(* IEC 61131-3 sources: IRIS-Project/LASAL CONTROL SOFTWARE/LasalProject_2025_09_12/Runtime/%LASALAPPDATA%/Runtime/Library/Loader/Source/code (part 4) *)

Find_sRam_I_END

END_FUNCTION // Find_sRam_I
#endif

FUNCTION GLOBAL Find_sRamEx
VAR_INPUT
	CRC32		: UDINT;
  bDontAdd : BOOL;
END_VAR
VAR_OUTPUT
	pRamAdr			: ^XramCell;
END_VAR
VAR
	pRamAdr_Kopie	: ^XramCell;
	udAllocated : UDINT;
	udLength : UDINT;
	RelAdress		: UDINT;
	pData : ^USINT;
	pData_Kopie : ^USINT;
	errCode : DINT;
	rc : DINT;
END_VAR

	IF fReorgSram THEN
		rc := LoadSramKopie(#errCode, 0, 0);
		IF rc <> 0 THEN
			// das Laden de SRAM Kopie hat nicht funktioniert
			fReorgSram := 0;
			DEBUGLOG2("%010d LoadSramKopie failed, rc=%d, errCode = 0x%X" , rc$UDINT, errCode$UDINT);
		END_IF;
	END_IF;

	IF fReorgSram THEN
		// in der Kopie suchen
		pRamAdr := Find_sRam_I(_S_RAM_Hptr_Kopie, CRC32);
	ELSE
		// im SRAM suchen
		pRamAdr := Find_sRam_I(_S_RAM_Hptr, CRC32);
	END_IF;

	IF pRamAdr = NIL THEN
		// nicht gefunden (weder im SRAM noch in der Kopie), neue Zelle anlegen
    if(bDontAdd = FALSE) then
  		nbrOfCells_notFound += 1;
  		pRamAdr := Add_sRam_I(CRC32);
    end_if;

	ELSIF fReorgSram THEN
		// in der Kopie gefunden, Zelle aus der Kopie ins SRAM kopieren
		nbrOfCells_foundInCopy += 1;

		pRamAdr_Kopie := pRamAdr;
		pRamAdr := Add_sRam_I(CRC32);
		IF pRamAdr THEN
			IF (pRamAdr_Kopie^.udType AND 16#3C000000) = IsXram THEN
				// RAMEX Zelle
 		     	udLength := pRamAdr_Kopie^.udData shr 16;
				// wenn die Länge der Daten > 0 ist, dann muss das RAMEX Objekt mit
				// den Daten aus der Kopie vorgeladen und für gültig erklärt werden
				IF udLength > 0 THEN
				 	RelAdress$UDINT:= (SRAM_GetMemory(udLength))$UDINT;
				 	// --- Speicher ist zugewiesen worden --
				 	If RelAdress <> 0 THEN
				   		GET_USED_S_RAM();
				   		udAllocated		      := SRAM_GET_ALLOCATED(udLength);
			  	   		pRAMadr^.udData$UDINT := (udLength shl 16) or (udAllocated and 16#ffff);
				   		pRAMadr^.udType 	  := RelAdress;
				   		pData				  := _S_RAM_Hptr^.DataStart+RelAdress;
				   		pData_Kopie			  := _S_RAM_Hptr_Kopie^.DataStart+(pRamAdr_Kopie^.udType and 16#00FF_ffff);
				   		_memcpy(pData, pData_Kopie, udLength);   // Speicher aus dem Inhalt aus der Kopie vorladen
		           		MakeRamExChk(pRAMadr);

				 	// -- Kein speicher verfügbar !!
				 	ELSE

						pRAMadr := NIL;

				 	END_IF;
				ELSE
	           		MakeRamExChk(pRAMadr);
				END_IF;
			ELSE
				// RAM Zelle
				pRamAdr^.udData := pRamAdr_Kopie^.udData;
				pRamAdr^.udChk := pRamAdr^.udData + CRC32;
				pRamAdr^.udType := 16#C0000000;    // ganz am ende machen wir uns gültig !
			END_IF;
		END_IF;
	ELSE
		nbrOfCells_foundInSram += 1;
	END_IF;

END_FUNCTION

FUNCTION GLOBAL Find_sRam
VAR_INPUT
	CRC32		: UDINT;
END_VAR
VAR_OUTPUT
	pRamAdr			: ^XramCell;
END_VAR

  pRamAdr := Find_sRamEx(CRC32, FALSE);

END_FUNCTION

////////////////////////////////////////////////////////////////////
//
//  Die IDEE:
//
//  LDRMEM => STRUCT
//
//  +----+-------------------------------+------------------------
//  |INFO| Allocation Table:             |
//  |MAT |   einzele Bits geben benutze  |   DATEN in 16-Byte Blöcken
//  |    |   Blöcke an                   |
//  +----+-------------------------------+------------------------
//
//  Allocation Table:
//  - jedes Bit kennzeichnet einen Block in den Daten
//  - ein 1er im Bit sagt aus, daß der entsprechende Block in den Daten frei ist
//  - das MSB zeigt auf den Block mit der höheren Adresse
//
//
////////////////////////////////////////////////////////////////////

FUNCTION SRAM_GetMemoryEx
VAR_INPUT
   length0  : UDINT;
   pGotMemory : ^BOOL;  // Da beim Returnwert 0 nicht unterschieden werden kann, ob
                        // der Offset 0 gemeint ist oder Out-Of-Memory, wird mit diesem
                        // Flag angezeigt, ob Speicher allokiert werden konnte.
END_VAR
VAR_OUTPUT
   ret0 : ^USINT;
END_VAR
VAR
   allocblocknum : UDINT;
   allocblocknumorg : UDINT;
   matsize  : UDINT;
   actblockcount : UDINT;
   actblocknum : UDINT;
   fbptr:^usint;
   startptr:^usint;
   fb, xfb : usint;
   bitcounter:usint;
   start:usint;
   startbit:usint;
   bytecounter:udint;
END_VAR

  pGotMemory^ := FALSE;
  ret0 := NIL; 	//#FA16122003
  if length0 = 0 then
    ret0 := NIL;
    return;
  end_if;

  allocblocknum := ((length0-1) / pLdrmem^.blocksize)+1; // Anzahl der erforderlichen Blöcke
  allocblocknumorg := allocblocknum;
  matsize := pLdrmem^.matsize; // Größe der MAT in Bytes
  actblockcount := 0;
  fbptr := #pLdrmem^.mat[0];
  fb := fbptr^;
  start := 1; // 1=suche ersten freien Block, 0=freier wurde Block gefunden
  bytecounter := 0;

  // Schleife, in der die MAT nach einem zusammengehörenden Bereich mit freien
  // Blöcken (=gesetzten Bits) durchsucht wird.
  while matsize do
    fb := fbptr^;
    if fb then
      // das aktuelle Byte in der MAT ist <>0, d.h. manche Blöcke sind frei
      if start = 0 then
        bytecounter += 1;
      end_if;

      // alle Bits des Bytes fb durchgehen
      bitcounter := 0;
      while bitcounter < 8 do
        xfb := fb and 1;
        fb  := fb shr 1;
        if xfb then
          // wir sind innerhalb des Bytes auf einen freien Block gestoßen
          if start then
            // es handelt sich um den ersten freien Block
            start := 0;
            startptr := fbptr;
            startbit := bitcounter;
            allocblocknum := allocblocknumorg;
            actblocknum := actblockcount;
            bytecounter := 0;
          end_if;
          allocblocknum -= 1;
          if allocblocknum = 0 then
            // es wurde ein zusammenhängender Bereich freier Blöcke gefunden
            ret0 := NIL + ((actblocknum * 8) + startbit) * pLdrmem^.blocksize;
            pGotMemory^ := TRUE;

            // es müssen jetzt noch die Bits in der MAT auf den Wert 'belegt'(=0) geändert werden
            if bytecounter = 0 then   // startbit and endbit same byte
              // auf fb wird jetzt eine Maske geschrieben, mit der dann die Bits auf 0 ausmaskiert werden können
              if startbit = bitcounter then   // only a block of 16 byte
                fb := not (1 shl bitcounter);
              else
                bitcounter := 7 - bitcounter;
                fb := ((16#FF shr startbit) and 16#FF) shl startbit; // Bits rechts von startbit werden auf 0 gesetzt
                fb := ((fb shl bitcounter) and 16#FF) shr bitcounter; // Bits links von bitcounter werden auf 0 gesetzt
                fb := not fb; // Wert invertieren, damit er als UND-Maske verwendet werden kann
              end_if;
              startptr^ := startptr^ and fb; // Bits mit der Maske auf 0 ausmaskieren
            else // 1 byte between start and end
              fb := ((16#FF shr startbit) and 16#FF) shl startbit; // Bits rechts von startbit werden auf 0 gesetzt
              fb := not fb; // Wert invertieren, damit er als UND-Maske verwendet werden kann
              startptr^ := startptr^ and fb; // Bits mit der Maske auf 0 ausmaskieren
              startptr += 1;
              if bytecounter then
                bytecounter -= 1;
                // die Bytes zwischen dem ersten und letzten werden zur Gänze auf 0 gesetzt
                while bytecounter do
                  startptr^ := 0;
                  startptr += 1;
                  bytecounter -= 1;
                end_while;
              end_if;
              bitcounter := 7 - bitcounter;
              fb := ((16#FF shl bitcounter) and 16#FF) shr bitcounter;// Bits links von bitcounter werden auf 0 gesetzt
              fb := not fb; // Wert invertieren, damit er als UND-Maske verwendet werden kann
              startptr^ := startptr^ and fb; // Bits mit der Maske auf 0 ausmaskieren
            end_if;

            // Fertig !
            return;

          end_if;
        else
          // wir sind innerhalb des Bytes auf einen belegten Block gestoßen
          start := 1;
        end_if;
        bitcounter += 1;
      end_while;
    else // if fb
      // das aktuelle Byte in der MAT ist 0, d.h. alle Blöcke sind belegt
      start := 1;
    end_if;
    actblockcount += 1;
    fbptr += 1;
    matsize -= 1;
  end_while;

END_FUNCTION

FUNCTION GLOBAL SRAM_GetMemory
VAR_INPUT
   length0  : UDINT;
END_VAR
VAR_OUTPUT
   ret0 : ^USINT;
END_VAR
VAR
	gotMemory : BOOL;
END_VAR

  ret0 := SRAM_GetMemoryEx(length0, #gotMemory);

END_FUNCTION

//---------------------------------------------
// Speicher Belegen
//---------------------------------------------
// es werden immer ganze blöcke vergeben
// -> Raladdr0 = Startadresse im s-Ram
// ->  length0 = Speicherlänge
//     #FA vorsicht die length hat 2 teile byte0/1 ist die allocated length
//                                         byte2/3 ist die used length
//										   also ein mask ist wichtig

// Wenn in length0 das oberste Bit gesetzt ist, dann wird vor dem Belegen geprüft,
// ob der gesamte Bereich frei ist. Wenn er nicht frei ist, dann wird auch nichts
// belegt.

//<-- 0 wenn ok

// diese Funktion wird nur beim Start verwendet um die bereits belegten RAMZellen zu markieren
// in Version alt 1 Bit sind 16 Byte
// in Version neu 1 Bit sind  4 Byte (der Rest der INFO steht im File beim C-IPC)
// abfrage über version die in den oberen 16 Bit von DataValid steht

FUNCTION SRAM_MarkMemory2
VAR_INPUT
   reladdr0 :^usint;
   length0  : UDINT;
END_VAR
VAR_OUTPUT
   ret0 : DINT;
END_VAR

    IF length0 AND 16#80000000 THEN
        // prüfen, ob der gesamte Bereich belegt ist
        length0 -= 16#80000000;
        ret0 := SRAM_FreeMarkMemory(reladdr0$UDINT, length0, 0, TRUE);
        IF ret0 <> 0 THEN
            RETURN;
        END_IF;
    END_IF;

    ret0 := SRAM_FreeMarkMemory(reladdr0$UDINT, length0, 1(*mark*), FALSE);

END_FUNCTION

#ifdef _LSL_TARGETARCH_ARM
FUNCTION GLOBAL SRAM_MarkMemory
VAR_INPUT
   reladdr0 :^usint;
   length0  : UDINT;
END_VAR
VAR_OUTPUT
   ret0 : DINT;
END_VAR

  ret0 := SRAM_MarkMemory2(reladdr0, length0);

END_FUNCTION
#else
FUNCTION AWL GLOBAL SRAM_MarkMemory
VAR_INPUT
   reladdr0 :^usint;
   length0  : UDINT;
END_VAR
VAR_OUTPUT
   ret0 : DINT;
END_VAR
    PUSHAD

    push      eax         //Result
    push.d    length0
    push.d    reladdr0

    call      SRAM_MarkMemory2

    add.esp   8
    pop.d     ret0        //Result

	POPAD

END_FUNCTION
#endif

#ifdef _LSL_TARGETARCH_ARM
FUNCTION GLOBAL SRAM_UnmarkMemory
VAR_INPUT
   reladdr0 :^usint;
   length0  : UDINT;
END_VAR
VAR_OUTPUT
   ret0 : DINT;
END_VAR

  ret0 := SRAM_FreeMarkMemory(reladdr0$UDINT, length0, 0(*0=Free Memory*), 0(*FALSE:ändern*));

END_FUNCTION
#else
FUNCTION AWL GLOBAL SRAM_UnmarkMemory
VAR_INPUT
   reladdr0 :^usint;
   length0  : UDINT;
END_VAR
VAR_OUTPUT
   ret0 : DINT;
END_VAR
    PUSHAD

    //#SR 16.12.2005
    push      eax         //Result
    push.d    0           //check
    push.d    0           //for unmark memory
    push.d    length0
    push.d    reladdr0

    call      SRAM_FreeMarkMemory

    add.esp   16
    pop.d     ret0        //Result

	POPAD

END_FUNCTION
#endif

//-------------------------------------------
//--- S-Ram Speicherverwaltung Initialisieren
//-------------------------------------------

// Hat a.m geprüft

FUNCTION GLOBAL SRAM_Startup
VAR_INPUT
   length0  : UDINT;
   clear0   : UDINT;
END_VAR
VAR_OUTPUT
   ret0 : DINT;
END_VAR
VAR
   matsize  : UDINT;
   memlength  : UDINT;
END_VAR

   ret0 := -1; // desciptior fehlerhaft, nichts gibts für die ramexerei

   // Größe der MAT ermitteln
   if !!isRamfileDatUsed | ((_S_RAM_Hptr^.DataValid SHR 16) < 2)  then
    matsize   := length0 / (CST_SRAM_BLOCKSIZE * 8); // anzahl der BitMarker
    memlength := matsize * (CST_SRAM_BLOCKSIZE * 8);
   else
    matsize   := 4 * length0 / (CST_SRAM_BLOCKSIZE * 8); // anzahl der BitMarker
    memlength := matsize * (CST_SRAM_BLOCKSIZE * 8) / 4;
   end_if;

   IF pLdrmem = NIL THEN
    // MAT neu allokieren
	// pr:
	//	In der Funktion SRAM_ClearMAT wird um ein DWORD mehr als matsize initialisiert,
	//  daher müssen 4 Bytes zusätlich allokiert werden. Den Grund für die zusätzlichen
	//	4 Bytes kenne ich nicht.
   	pLdrmem := _alloc_resize_LDR(MAT_INFO_TYPE.mat + matsize + 4)$^MAT_INFO_TYPE;
   ELSIF pLdrmem^.matsize <> matsize THEN
    // Größe der MAT ändern
   	pLdrmem := _realloc_LDR(pLdrmem, MAT_INFO_TYPE.mat + matsize + 4)$^MAT_INFO_TYPE;
   END_IF;

   IF pLdrmem = NIL THEN
    ret0 := -1;
    RETURN;
   END_IF;

   pLdrmem^.memlength := memlength;
   pLdrmem^.matsize   := matsize;
   if !!isRamfileDatUsed | ((_S_RAM_Hptr^.DataValid SHR 16) < 2)  then
	pLdrmem^.blocksize := CST_SRAM_BLOCKSIZE;
   else
	pLdrmem^.blocksize := CST_SRAM_BLOCKSIZE_NEW;
   end_if;

   if clear0 then
    SRAM_ClearMAT();
   end_if;

   ret0 := 0; // alles ist gut, daher probieren mal eine kleine ramexerei
END_FUNCTION

//---------------------------------------------
// -- ALLE Blockmarker mit 1 auf "leer" setzen
//---------------------------------------------
#ifdef _LSL_TARGETARCH_ARM
FUNCTION GLOBAL SRAM_ClearMAT

  _memset(#pLdrmem^.mat[0], 16#ff, pLdrmem^.matsize);

END_FUNCTION
#else
FUNCTION AWL GLOBAL SRAM_ClearMAT

		l.ecx		pLdrmem
   		l.ecx		(ecx + MAT_INFO_TYPE.matsize)
		shr.ecx		2				// /4
		jecxz		SRAM_ClearMATRet

		// pr: wozu das ???
		// ** Fehler IPC 300 **     // es wird mehr eigetragen wie vorhandener speicher
		inc			ecx				// wegen IPC 300 sonst werden die Daten nicht gespeichert

		l.edi		pLdrmem
		add.edi		MAT_INFO_TYPE.mat
		l.eax		16#ffffffff
		rep
		stosd
SRAM_ClearMATRet
END_FUNCTION
#endif

//-----------------------------------
// Liefert Die Belegte Speichergrösse (bezogen auf speicherstart)
//-----------------------------------
FUNCTION GLOBAL SRAM_GetLastAddr
VAR_OUTPUT
   ret0 : UDINT;
END_VAR
VAR
   Lng: UDINT;
   size:udint;
   Muster : BSINT;
   fbptr : ^bsint;
END_VAR
   fbptr := #pLdrmem^.mat[pLdrmem^.matsize-1];  // in letzet eintrag im array

   Lng    := pLdrmem^.memlength;				// beginn bei voller belegung
   size   := pLdrmem^.matsize;

   while size do
      if fbptr^ <> 16#FF then     			// erster freier platz wenn nicht auf FF
		 Muster:=fbptr^ $bsint;
		 While Muster do
           Lng-=pLdrmem^.blocksize;
		   muster := muster SHL 1;
		 end_while;
		 Goto  LastAdrEnde;

      end_if;
      fbptr -= 1;
	  size -= 1;
	  Lng-= pLdrmem^.blocksize*8;
   end_while;

LastAdrEnde:
   ret0 := Lng;
END_FUNCTION

(*
    Markiert im Sram in der MAT einen Bereich als frei oder belegt oder
    prüft ob der Bereich vollständig frei oder vollständig belegt ist.
*)
FUNCTION SRAM_FreeMarkMemory
VAR_INPUT
    reladdr0 : UDINT;
    length0  : UDINT;
    mode0    : UDINT;        //0=Free Memory, 1=Mark Memory
    check0   : BOOL;         //FALSE:ändern, TRUE:nur prüfen
END_VAR
VAR_OUTPUT
    ret0 : DINT;
END_VAR
VAR
    startBit : UDINT;
    endBit : UDINT;
    curBit : UDINT;
    ofs : UDINT;
    pMat : ^USINT;
    matVal : USINT;
END_VAR

    ret0 := 0;

    IF ((reladdr0 + length0) > pLdrmem^.memlength) | (length0 = 0) THEN
        // Der angegebene Bereich liegt ausserhalb der Grenzen oder die Länge ist 0 -> Fehler zurückgeben
        ret0 := -1;
        RETURN;
    END_IF;

    startBit := reladdr0 / pLdrmem^.blocksize;
    endBit := (reladdr0 + length0 - 1) / pLdrmem^.blocksize;
    IF mode0 = 0 THEN
        matVal := 0xFF;
    ELSE
        matVal := 0x00;
    END_IF;

    curBit := startBit;
    pMat := #pLdrmem^.mat[curBit / 8];
    WHILE curBit <= endBit DO
        ofs := curBit MOD 8;
        IF (ofs = 0) & ((endBit - curBit) >= 8) THEN
            // Wir befinden uns auf einer Byte-Grenze daher können alle 8 Bits
            // des MAT-Bytes auf einmal behandelt werden.
            IF check0 THEN
                // nur prüfen
                IF pMat^ <> matVal THEN
                    ret0 := -1;
                    RETURN;
                END_IF;
            ELSE
                // ändern
                pMat^ := matVal;
            END_IF;

            curBit += 8;
            pMat += 1;
        ELSE
            // Wir befinden uns mitten im Byte. Die Bits müssen einzeln behandelt werden.
            IF check0 THEN
                // nur prüfen
                IF mode0 = 0 THEN
                    IF (pMat^ AND (1 SHL ofs)$USINT) = 0 THEN
                        ret0 := -1;
                        RETURN;
                    END_IF;
                ELSE
                    IF (pMat^ AND (1 SHL ofs)$USINT) <> 0 THEN
                        ret0 := -1;
                        RETURN;
                    END_IF;
                END_IF;
            ELSE
                // ändern
                IF mode0 = 0 THEN
                    pMat^ := pMat^ OR (1 SHL ofs)$USINT;
                ELSE
                    pMat^ := pMat^ AND NOT (1 SHL ofs)$USINT;
                END_IF;
            END_IF;

            curBit += 1;
            IF (curBit MOD 8) = 0 THEN
                pMat += 1;
            END_IF;
        END_IF;
    END_WHILE;

END_FUNCTION

#ifdef LDR_RETSVR
FUNCTION GLOBAL GetNbrNotFound
VAR_OUTPUT
  ret0 : udint;
END_VAR

  ret0 := nbrOfCells_notFound;

END_FUNCTION

// ein neues File muss erstellt werden
FUNCTION NewRetainSvrFile
	VAR_INPUT
		usProbe 	: usint;
	END_VAR
  VAR_OUTPUT
    ok : dint;
  END_VAR
  var
    pRead : ^MRAM_DESCR;
    pData : ^MRAM_DESCR;
  end_var

  // Schreib-/Lesebuffer
  pData := _alloc_resize_LDR( sizeof( MRAM_DESCR ) * 2 )$^MRAM_DESCR;
  pRead := pData + sizeof( MRAM_DESCR );

  if( pData <> NIL )then

    // einen gültigen Header erzeugen
    _memset( pData, 16#00, sizeof( MRAM_DESCR ) * 2 );
    pData^.version     := 0;
    pData^.DataStart   := 20;
    pData^.DataLength  := -1$udint; //wir sehen mal keine Längenbegrenzung vor
    pData^.UsedData    := 20;
    pData^.DataValid   := 1;

    if( FileWrite( hLDR_remSvr, pData, sizeof( MRAM_DESCR ) ) = sizeof( MRAM_DESCR ) )then

      // schauen, ob das Filesystem auch beschreibbar ist
      if( OS_FILE_SEEK( hLDR_remSvr, 0, FILE_BEGIN ) = 0 )then
        if( OS_FILE_READ( hLDR_remSvr, pRead, sizeof( MRAM_DESCR ) ) = sizeof( MRAM_DESCR ) )then
          if( _memcmp( pData, pRead, sizeof( MRAM_DESCR ) ) = 0 )then

            ok := 1;

            //nur Probe, dann wieder schließen
            if( usProbe )then
              OS_FILE_CLOSE( hLDR_remSvr );
              OS_FILE_DELETE( LDR_RETENTIVE_SVRFILENAME );
              hLDR_remSvr := 0;
            else
            // sonst den Zeiger wieder auf den Fileanfang
              OS_FILE_SEEK( hLDR_remSvr, 0, FILE_BEGIN );
            end_if;
          end_if;
        end_if;
      end_if;
    end_if;
    _free( pData );
  end_if;

END_FUNCTION

// Initialisiert das File zum Speichern der remanenten Server
// > usProbe: 1..nur schauen, obs prinzipiell geht
//            0..das File auch gleich öffnen (offen lassen)
FUNCTION GLOBAL InitRetainSvrFile
	VAR_INPUT
		usProbe 	: usint;
	END_VAR
	VAR_OUTPUT
		ok 	: DINT;
	END_VAR

  if( hLDR_remSvr <> 0 )then
    ok := 1;
    return;
  end_if;

  ok := 0;

  //existiert das File
  hLDR_remSvr := OS_FILE_OPEN( LDR_RETENTIVE_SVRFILENAME, 2, ATT_OPEN_SHARED or ATT_COMMITTED);

  if( hLDR_remSvr >= 0 )then

    //Fileinhalt checken
    if( LoadSramKopie( NIL, hLDR_remSvr, usProbe ) = 0 )then
      ok := 1;
    else
      DEBUGLOG0("%010d-InitRetainSvrFile: file corrupted. Stored in retsvr.err and generated a new one!");
      TRACE_ERR("Error in RetSvrFile, see c:\sysmsg\event19.log");
      LSLCLI_LoaderTracePrint("Error in RetSvrFile, see c:\sysmsg\event19.log", 12);
      OS_FILE_CLOSE( hLDR_remSvr );
      OS_FILE_RENAME( LDR_RETENTIVE_SVRFILENAME, LDR_RETENTIVE_SVRFILENAME_ERR );
      hLDR_remSvr := OS_FILE_OPEN( LDR_RETENTIVE_SVRFILENAME, 2, ATT_OPEN_SHARED or ATT_CREATE_ALWAYS or ATT_COMMITTED);
      if( hLDR_remSvr >= 0 )then
        //Schreib/Lesetest
        ok := NewRetainSvrFile( usProbe );
      end_if;
    end_if;

    //nur Probe, dann wieder schließen
    if( ( usProbe <> 0 ) | ( ok = 0 ) )then
      OS_FILE_CLOSE( hLDR_remSvr );
      hLDR_remSvr := 0;
    end_if;
  else
  //nein, dann anlegen und testen
    hLDR_remSvr := OS_FILE_OPEN( LDR_RETENTIVE_SVRFILENAME, 2, ATT_OPEN_SHARED or ATT_CREATE_ALWAYS or ATT_COMMITTED);
    if( hLDR_remSvr >= 0 )then
      DEBUGLOG0("%010d-InitRetainSvrFile: created new retsvr.dat");

      //Schreib/Lesetest
      ok := NewRetainSvrFile( usProbe );
      if( ( usProbe <> 0 ) | ( ok = 0 ) )then
        OS_FILE_CLOSE( hLDR_remSvr );
        hLDR_remSvr := 0;
      end_if;
    else
      hLDR_remSvr := 0;
    end_if;
  end_if;

END_FUNCTION

// Gibt den temporären Speicher frei
FUNCTION GLOBAL FreeMemoryRetainSvrFile
var
  a : ^MRAM_DESCR;
end_var
  // den Buffer vor dem reorg brauchen wir gar nicht mehr
  if( _S_RAM_Hptr_File <> NIL )then
    _free( _S_RAM_Hptr_File );
    _S_RAM_Hptr_File := NIL;

    // der reorganisiserte Bufer landet im File
    a := _S_RAM_Hptr_File_New;
    if( _S_RAM_Hptr_File_New <> NIL )then
      if( OS_FILE_SEEK( hLDR_remSvr, 0, FILE_BEGIN ) = 0 )then
        if( FileWrite( hLDR_remSvr, _S_RAM_Hptr_File_New, _S_RAM_Hptr_File_New^.UsedData )$UDINT = _S_RAM_Hptr_File_New^.UsedData )then

          // und das File schneiden wir auf die benötigte Länge zu
          OS_FILE_TRUNCATE( hLDR_remSvr );
          OS_FILE_SEEK( hLDR_remSvr, 0, FILE_BEGIN );
        else
          DEBUGLOG0("%010d-FreeMemoryRetainSvrFile: Cannot reorg.!");
        end_if;
      else
        DEBUGLOG0("%010d-FreeMemoryRetainSvrFile: Cannot reorg.!");
      end_if;
      _free( _S_RAM_Hptr_File_New );
      _S_RAM_Hptr_File_New := NIL;
    end_if;
  end_if;

END_FUNCTION

(*
  Hängt eine ASYNC_FILE_STATE Datenstruktur ans Ende der verketteten Liste an.
*)
FUNCTION AppendAsyncState
VAR_INPUT
  pAsyncState : ^RetSvrFile::ASYNC_FILE_STATE;
END_VAR

  IF pAsyncState^.pNext <> NIL THEN
    // Dieser Zustand darf nie eintreten. Wenn doch, dann Excepion auslösen
    (0$^UDINT)^ := 0;
  END_IF;

  IF pLastAsyncState = NIL THEN
    IF pFirstAsyncState <> NIL THEN
      // Dieser Zustand darf nie eintreten. Wenn doch, dann Excepion auslösen
      (0$^UDINT)^ := 0;
    END_IF;
    pFirstAsyncState := pAsyncState;
    pLastAsyncState := pAsyncState;
  ELSE
    pLastAsyncState^.pNext := pAsyncState;
    pLastAsyncState := pAsyncState;
  END_IF;

  nAsyncStateObjs += 1;

END_FUNCTION

(*
  Entfernt eine ASYNC_FILE_STATE Datenstruktur aus der verketteten Liste.
*)
FUNCTION RemoveAsyncState
VAR_INPUT
  pPrev : ^RetSvrFile::ASYNC_FILE_STATE;
  pAsyncState : ^RetSvrFile::ASYNC_FILE_STATE;
END_VAR

  IF pPrev = NIL THEN
    // es wird das Element am Anfang entfernt
    pFirstAsyncState := pAsyncState^.pNext;
  ELSE
    // es wird ein Element nach dem Anfang entfernt
    pPrev^.pNext := pAsyncState^.pNext;
  END_IF;
  IF pAsyncState = pLastAsyncState THEN
    // es wird das Element am Ende entfernt
    pLastAsyncState := pPrev;
  END_IF;

  pAsyncState^.pNext := NIL;

  nAsyncStateObjs -= 1;

END_FUNCTION

FUNCTION Get_ITASK_Version
VAR_OUTPUT
	version : UDINT;
END_VAR

  // Anm.: Beim Salamander darf das udVersion Element aus der LSL_ITASK Struktur
  // (Makro OS_ITASK_VERSION) erst ab 09.03.080 interpretiert werden, weil sonst
  // keine Versionsnummer dahintersteckt, sondern ein Funktionszeiger auf eine Dummy-Funktion.
  IF _RtOSVersion < 16#9000 | _RtOSVersion >= 16#9350 THEN
    version := OS_ITASK_VERSION;
  ELSE
    version := 0;
  END_IF;

END_FUNCTION

(*
  Liefert die Info, ob das OS versucht, die Applikation zu stoppen
*)
FUNCTION ITASK_IS_STOPPING
VAR_OUTPUT
  is_stopping : UDINT;
END_VAR

  IF Get_ITASK_Version() >= 0x11 THEN
    is_stopping := OS_ITASK_IS_STOPPING();
  ELSE
    is_stopping := 0;
  END_IF;

END_FUNCTION

(*
  Inkrementiert oder dekrementiert den StopWait Zähler.
  Wenn dieser >0 ist dann wartet das OS beim Stoppen der Applikation, bis dieser
  Zähler auf 0 geht. Die Applikation kann damit das Stoppen der Applikation
  verzögern bis z,B. alle Retentive File Server geschrieben sind.
*)
FUNCTION ITASK_SET_STOPWAIT_CNTR
VAR_INPUT
  inc_dec : DINT;
END_VAR

  IF Get_ITASK_Version() >= 0x11 THEN
    OS_ITASK_SET_STOPWAIT_CNTR(inc_dec);
  END_IF;

END_FUNCTION

(*
  Asynchrone Version von RetSvrFileWrite.

  Diese Funktion wird von einem RetSvrFile Objekt aufgerufen, wenn die XRamCell Struktur des
  Objekts ins remanente File geschrieben werden soll. Das Schreiben erfolgt asynchron.
  Der Request wird in die Liste pFirstAsyncState eingetragen. Diese Liste wird in der
  zyklischen Loaderfunktion ProcessAsyncFileObjects abgearbeitet.
*)
FUNCTION GLOBAL RetSvrFileWrite_A
VAR_INPUT
  pAsyncState : ^RetSvrFile::ASYNC_FILE_STATE;  // Zeiger auf eine bereits initialisierte ASYNC_FILE_STATE Struktur
END_VAR
VAR_OUTPUT
  ret0 : dint;
END_VAR
VAR
	pCell : ^XRamCell;
END_VAR

  ret0 := -1;

  IF processAsyncFileError < 0 THEN
    return;
  END_IF;

  IF ITASK_IS_STOPPING() THEN
    // Wenn das Betriebsystem gerade versucht, die Applikation zu stoppen,
    // wird kein neuer Schreibrequest angenommen.
    RETURN;
  END_IF;

  pCell := #pAsyncState^.XRamAddr;

  // wenn wir das Projekt grad hochfahren, dann darf nichts in das File geschrieben werden!
  // das landet (vorerst) alles im Buffer und wird beim Reorg geschrieben
  if( _S_RAM_Hptr_File_New = NIL )then

    // existiert das Handle?
    if( hLDR_remSvr <> NIL )then
      OS_MT_Wait(hMemMutex);
      IF pAsyncState^.state = 0 THEN
        // pAsyncState an die Liste der AsyncState Objekte hinten anhängen
        AppendAsyncState(pAsyncState);
      END_IF;
      pAsyncState^.state := pAsyncState^.state OR 1; // State 1 bedeutet, dass pDataObj^ geschrieben werden muss
      IF !!AsnycFileOperationInProgress THEN
        // Wird haben in einen Zustand gewechselt, in dem Daten gespeichert sind,
        // die erst geschrieben werden müssen. Dem Betriebssystem wird das mit dem
        // Aufruf der ITASK_SET_STOPWAIT_CNTR(1) mitgeteilt.
        ITASK_SET_STOPWAIT_CNTR(1);
      END_IF;
      AsnycFileOperationInProgress := TRUE;
      OS_MT_Signal(hMemMutex);
    end_if;

  else
    pCell^.udData := pAsyncState^.pDataObj^;
    _memcpy( _S_RAM_Hptr_File_New + pCell^.udType, pCell, sizeof( XRamCell ) );
  end_if;

  ret0 := 0;

END_FUNCTION

(*
  Bearbeitet eine asynchronene File Datenstruktur eines RetSvrFile Objekts.

  Hier wird das asynchrone Fileschreiben angestossen und überwacht. Sobale eine asynchrone Fileoperation
  fertig ist, wird das Element state der Struktur auf 0 gesetzt.

  Return:
    1 wenn kein schwerwiegender Fehler aufgetreten ist und die aüssere Schleife abgebrochen werden
      soll
    0 wenn kein schwerwiegender Fehler aufgetreten ist
   <0 wenn ein schwerwiegender Fehler aufgetreten ist, bei dem man annehmen muss, dass das File korrupt ist
        und deswegen auf ungültig gesetzt werden muss.
*)
FUNCTION ProcessOneAsyncFileObject
VAR_INPUT
	pAsyncState : ^RetSvrFile::ASYNC_FILE_STATE;
END_VAR
VAR_OUTPUT
  result : DINT;
END_VAR
VAR
	pCell : ^XRamCell;
  rc : DINT;
  requestResult : DINT;
  itoa_buf : ARRAY[0..20] OF CHAR;
END_VAR

  result := 0;

  IF pAsyncState^.state = 1 THEN
    IF (_rtosversion < (16#1200 + 93)) & (nAsyncStateReqs > 0) THEN
      // Bei einer OS Version < 1.2.93 kommte es zu einem Fehler, wenn die Async-Mailbox voll wird,
      // daher wird in so einem Fall nur dann etwas neues in die Mailbox gestellt, wenn gerade
      // kein Request unterwegs ist (Anzahl der anstehenden Requests steht in nAsyncStateReqs)
      result := 1;
      RETURN;
    END_IF;
    pCell := #pAsyncState^.XRamAddr;
    rc := OS_FILE_SEEK_AV1(Async0:=1, handle0:=hLDR_remSvr, offset0:=pCell^.udType$DINT, fromwhere0:=FILE_BEGIN);
#ifdef TEST_RETSVRFILE  // Code kann für Testzwecke aktiviert werden
    IF simuFSeekA_error <> 0 THEN
      rc := simuFSeekA_error;
    END_IF;
#endif
    IF rc >= 0 THEN
      // Request fürs Positionieren wurde angenommen

      // Daten in die XRamCell übernehmen
      pCell^.udData := pAsyncState^.pDataObj^;
      // asynchrones FileWrite anstossen
      rc := OS_FILE_WRITE_AV1(Async0:=1, fhandle0:=hLDR_remSvr, buffer0:=pCell, length0:=sizeof(XRamCell));
#ifdef TEST_RETSVRFILE  // Code kann für Testzwecke aktiviert werden
      IF simuFWriteA_error <> 0 THEN
        rc := simuFWriteA_error;
      END_IF;
#endif
      IF rc >= 0 THEN
        // Request konnte abgesetzt werden -> Request-Handle merken und Status aktualisieren
        pAsyncState^.hRequest := rc;
        pAsyncState^.state := 2;
        nAsyncStateReqs += 1;
      ELSIF rc = -200 THEN // -200=Mailbox voll
        result := 1; // Bearbeitung der restlichen Listeneinträge kann entfallen
        RETURN;
      ELSE
      	_itoa(rc$UDINT, #itoa_buf[0]);
        TRACE0_ERR("ERROR in ProcessOneAsyncFileObject: OS_FILE_WRITE_AV1 failed, {0}", #itoa_buf[0]);
      END_IF;
    ELSIF rc = -200 THEN // -200=Mailbox voll
      result := 1; // Bearbeitung der restlichen Listeneinträge kann entfallen
      RETURN;
    ELSE
      // SA33172,DS2528:
      // In diesem Fall (OS_FILE_SEEK_AV1 hat einen Fehler <> -200 geliefert), wird die
      // Bearbeitung der restlichen Listeneinträge abgebrochen, weil sonst bei einem
      // permanenten Fehler auf der SD-Karte die CPU-Belastung sehr hoch werden würde.
      result := 1;
    	_itoa(rc$UDINT, #itoa_buf[0]);
      TRACE0_ERR("ERROR in ProcessOneAsyncFileObject: OS_FILE_SEEK_AV1 failed, {0}", #itoa_buf[0]);
    END_IF;
  END_IF;

  IF pAsyncState^.state > 1 THEN
    rc := OS_FILE_GETASYNCSTATE(ID:=pAsyncState^.hRequest$UDINT, Erg:=#requestResult);
    IF rc >= 0 THEN
      // Request ist abgeschlossen -> Ergebnis der Fileoperation prüfen und Status aktualisieren
#ifdef TEST_RETSVRFILE  // Code kann für Testzwecke aktiviert werden
      IF simuFReq_error <> 0 THEN
        requestResult := simuFReq_error;
      END_IF;
#endif
      IF requestResult < 0 THEN
        result := requestResult;
      END_IF;
      pAsyncState^.state := pAsyncState^.state AND (NOT 2);
      pAsyncState^.wrCnt += 1;
      nAsyncStateReqs -= 1;
      IF pAsyncState^.state = 1 THEN
        (* Wir sind jetzt in der Situation dass während der asynchronen Fileoperation wieder das
           dData des RetSvrFile Objekts beschrieben worden ist. Wenn man jetzt nichts unternimmt,
           dann könnte für dieses Objekt beim nächsten Durchlauf wieder ein Request abgesetzt werden.
           Wenn sich dieses Spielchen ständig wiederholt, dann könnten andere Objekte mit Status 1,
           die sich in der Liste weiter hinten befinden, möglicherweise nie gestartet werden.
           Um das zu verhindern, sollte diese Objekt aus der Liste entfernt und hinten wieder
           angehängt werden. Das muss vom Aufrufer erledigt werden und damit er weiss dass er das
           machen soll, wird der state auf den temporären Wert 4 gesetzt.
         *)
         pAsyncState^.state := 4;
      END_IF;
    ELSIF rc = RT_NOT_STARTED | rc = RT_IN_PROGRESS THEN
      result := 1; // Bearbeitung der restlichen Listeneinträge kann entfallen
      RETURN;
    ELSE
    	_itoa(rc$UDINT, #itoa_buf[0]);
      TRACE0_ERR("ERROR in ProcessOneAsyncFileObject: OS_FILE_GETASYNCSTATE failed, {0}", #itoa_buf[0]);
    END_IF;
  END_IF;

END_FUNCTION

(*
  Bearbeitet alle Elemente in der Liste der asynchronen File Datenstrukturen von RetSvrFile Objekten.

  Für jedes Element wird ProcessOneAsyncFileObject aufgerufen und wenn dann angezeigt wird, dass die
  asynchrone Fileoperation fertig ist, wird das aktuelle Element aus der Liste entfernt.
*)
FUNCTION GLOBAL ProcessAsyncFileObjects
VAR
	pAsyncState : ^RetSvrFile::ASYNC_FILE_STATE;
	pPrev : ^RetSvrFile::ASYNC_FILE_STATE;
	pNext : ^RetSvrFile::ASYNC_FILE_STATE;
  rc : DINT;
  validFlag : UDINT;
END_VAR

  IF processAsyncFileError < 0 THEN
    return;
  END_IF;

  rc := 16#12345678;

  // Mit dieser Abfrage wird der OVerhead von OS_MT_Wait/OS_MT_Signal vermieden,
  // wenn nichts abzuarbeiten ist.
  IF pFirstAsyncState <> NIL THEN
    OS_MT_Wait(hMemMutex);
    pPrev := NIL;
    pAsyncState := pFirstAsyncState;
    WHILE pAsyncState <> NIL DO
      IF pAsyncState^.state = 0 THEN
        // Dieser Zustand darf nie eintreten. Wenn doch, dann Excepion auslösen
        (0$^UDINT)^ := 0;
      END_IF;

      rc := ProcessOneAsyncFileObject(pAsyncState);
      IF rc < 0 THEN
        // schwerweigender Fehler, File ist möglicherweise korrupt
        // -> File als ungültig markieren, Fehlerflag setzen
        validFlag := 0;
        OS_FILE_SEEK( hLDR_remSvr, MRAM_DESCR.DataValid, FILE_BEGIN );
        FileWrite( hLDR_remSvr, #validFlag$^void, sizeof( MRAM_DESCR.DataValid ) );
        processAsyncFileError := rc;
      END_IF;
      IF rc = 1 THEN
        EXIT;
      END_IF;

      pNext := pAsyncState^.pNext;
      IF pAsyncState^.state = 0 THEN
        // state 0: Request wurde beendet -> Objekt entfernen
        RemoveAsyncState(pPrev, pAsyncState);
      ELSIF pAsyncState^.state = 4 THEN
        // state 4: Request wurde beendet, dData wurde aber zwischenzeitlich wieder geändert
        //  -> Objekt entfernen und hinten wieder anhängen
        RemoveAsyncState(pPrev, pAsyncState);
        pAsyncState^.state := 1;
        AppendAsyncState(pAsyncState);
      ELSE
        pPrev := pAsyncState;
      END_IF;
      pAsyncState := pNext;
    END_WHILE;
    OS_MT_Signal(hMemMutex);
  END_IF;

  if((rc = 0) | (rc = 16#12345678)) then
    OS_MT_Wait(hMemMutex);
    IF AsnycFileOperationInProgress THEN
      // Wird haben den Zustand verlassen, in dem Daten gespeichert sind,
      // die erst geschrieben werden müssen. Dem Betriebssystem wird das mit dem
      // Aufruf der ITASK_SET_STOPWAIT_CNTR(-1) mitgeteilt.
      ITASK_SET_STOPWAIT_CNTR(-1);
    END_IF;
    AsnycFileOperationInProgress := FALSE;
    OS_MT_Signal(hMemMutex);
  end_if;

END_FUNCTION

FUNCTION GLOBAL LDR_IsAsnycFileOperationInProgress
VAR_OUTPUT
  ret   : BOOL;
END_VAR

  ret := AsnycFileOperationInProgress;
END_FUNCTION

FUNCTION GLOBAL LDR_HasSram
VAR_OUTPUT
  ret   : BOOL;
END_VAR

  ret := hasSram;
END_FUNCTION

#if 0
FUNCTION GLOBAL RetSvrFileWrite
VAR_INPUT
  pCell : ^XRamCell;
END_VAR
VAR_OUTPUT
  ret0 : dint;
END_VAR

  ret0 := -1;

  // wenn wir das Projekt grad hochfahren, dann darf nichts in das File geschrieben werden!
  // das landet (vorerst) alles im Buffer und wird beim Reorg geschrieben
  if( _S_RAM_Hptr_File_New = NIL )then

    // existiert das Handle?
    if( hLDR_remSvr <> NIL )then

      // auf die gewünschte Zelle positionieren
      if( OS_FILE_SEEK( hLDR_remSvr, pCell^.udType, FILE_BEGIN ) = pCell^.udType )then
        pCell^.udChk := pCell^.udData;

        // und reinschreiben
        if( OS_FILE_WRITE( hLDR_remSvr, pCell, sizeof( XRamCell ) ) = sizeof( XRamCell ) )then
          ret0 := 0;
        else
          ret0 := -2;
        end_if;
      else
        ret0 := -2;
      end_if;
    end_if;

    // Positionieren oder Schreiben hat nicht hingehaun -> File ist korrupt!
    if( ret0 = -2 )then
      OS_FILE_SEEK( hLDR_remSvr, MRAM_DESCR.DataValid, FILE_BEGIN );
      ret0 := 0;
      OS_FILE_WRITE( hLDR_remSvr, #ret0$^void, sizeof( MRAM_DESCR.DataValid ) );
      ret0 := -2;
    end_if;
  else
    _memcpy( _S_RAM_Hptr_File_New + pCell^.udType, pCell, sizeof( XRamCell ) );
  end_if;

END_FUNCTION
#endif

#endif // LDR_RETSVR
